Universal Robots PolyScope program: P1140 INVITE.urp

Program P1140 INVITE (installation=default directory=/programs/02 Main Routines createdIn=5.10.1 lastSavedIn=5.19.0 robotSerialNumber=20245590068)
Calibrated DH parameters: a=[0.00013, -0.03651, -0.389144, 0.000102, 0.000008, 0]; d=[0.162613, 192.230671, -179.915756, -12.181517, 0.099698, 0.099535]; alpha=[1.57038, 0.002205, 0.004138, 1.570804, -1.571025, 0]; deltaTheta=[-0.000001, 1.484886, 4.928506, -0.130209, 0, 0]
InitVariablesNode variables(variable(name=AMR_Position, expression=struct(position_identifier=0, x1=0, x2=0, y1=0, y2=0, theta1=0, theta2=0)), variable(name=CAM_Pose, expression=p[0,0,0,0,0,0]), variable(name=CAM_Relation, expression=""), variable(name=CMD_Abort, expression=False), variable(name=CMD_Clear, expression=False), variable(name=CMD_Reset, expression=False), variable(name=CMD_Start, expression=False), variable(name=CMD_Suspend, expression=False), variable(name=CMD_Unhold, expression=False), variable(name=CMD_Unsuspend, expression=False), variable(name=CNT_Rack_Output, expression=0), variable(name=FNC_Freedrive, expression=False), variable(name=PRC_TubCounter, expression=0), variable(name=PRC_TubNumber, expression=0), variable(name=STP, expression=0), variable(name=TMR_Barcode, expression=0), variable(name=easyPickCount, expression=0), variable(name=easyPickCount_5, expression=0), variable(name=easyPickNoObj, expression=0), variable(name=easyPickNoObj_5, expression=0), variable(name=easyPickParts, expression=0), variable(name=easyPickParts_5, expression=0))
BeforeStart
  Folder Scripts [hidden by the author, left out]
  Folder BeforeStarts [hidden by the author, left out]
Robot Program (runOnlyOnce=false)
  Folder MAIN [hidden by the author, left out]
SubProgram -> Sub_Vision_V18
SubProgram  [hidden by the author, left out]
SubProgram  [hidden by the author, left out]
